// Mitsubishi GX Works2 project: Practica1   PLC: FX3G

PROGRAM MAIN
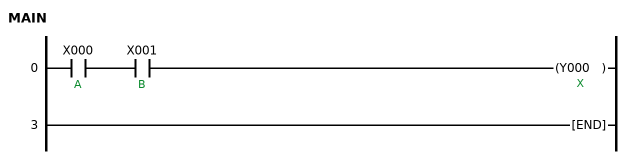
0     LD      X000  ; A
      AND     X001  ; B
      OUT     Y000  ; X
3     END
END_PROGRAM
